(* IEC 61131-3 sources: SRCI_CLIENT_PLC/RobotLibrary/Library/Enumerations/Level, 5 files *)

(* ---- LogLevel.st ---- *)
{attribute 'qualified_only'}
// -------------------------------------------------------------------------
//  SRCI Robot Library
// -------------------------------------------------------------------------
//
//  Object:      LogLevel
//  Author:      Thorsten Brach
//  Date:        2024-06-01
//
//  Description:
//
//
//  Copyright:
//    (C) 2024 Thorsten Brach. All rights reserved
//             Licensed under the MIT License.
//
//  Disclaimer:
//    This project is provided without any guarantee and can be used for
//    private and commercial purposes. Any use is at the user’s
//    own risk and responsibility.
//
// -------------------------------------------------------------------------
// ST-FIX W02: no attribute 'to_string' - LogLevel is an alias of Severity, the attribute is only valid for enumerations
TYPE LogLevel : Severity; END_TYPE

(* ---- LogLevelEnum.st ---- *)
TYPE LogLevelEnum : LogLevel; END_TYPE

(* ---- MessageLevel.st ---- *)
{attribute 'qualified_only'}
{attribute 'to_string'}
// -------------------------------------------------------------------------
//  SRCI Robot Library
// -------------------------------------------------------------------------
//
//  Object:      MessageLevel
//  Author:      Thorsten Brach
//  Date:        2024-06-01
//
//  Description:
//
//
//  Copyright:
//    (C) 2024 Thorsten Brach. All rights reserved
//             Licensed under the MIT License.
//
//  Disclaimer:
//    This project is provided without any guarantee and can be used for
//    private and commercial purposes. Any use is at the user’s
//    own risk and responsibility.
//
// -------------------------------------------------------------------------
TYPE MessageLevel :
(
  /// Debugging messages, Informative messages, Warning messages, Error messages, Fatal error messages
  DEBUG := 4,
  /// Informative messages, Warning messages, Error messages, Fatal error messages
  INFO := 5,
  /// Warning messages, Error messages, Fatal error messages
  WARNING := 20,
  /// Error messages, Fatal error messages
  ERROR := 28
)USINT;
END_TYPE

(* ---- MessageLevelEnum.st ---- *)
TYPE MessageLevelEnum : MessageLevel; END_TYPE

(* ---- PriorityLevel.st ---- *)
{attribute 'qualified_only'}
{attribute 'to_string'}
// -------------------------------------------------------------------------
//  SRCI Robot Library
// -------------------------------------------------------------------------
//
//  Object:      PriorityLevel
//  Author:      Thorsten Brach
//  Date:        2024-06-01
//
//  Description:
//
//
//  Copyright:
//    (C) 2024 Thorsten Brach. All rights reserved
//             Licensed under the MIT License.
//
//  Disclaimer:
//    This project is provided without any guarantee and can be used for
//    private and commercial purposes. Any use is at the user’s
//    own risk and responsibility.
//
// -------------------------------------------------------------------------
TYPE PriorityLevel :
(
  /// priority level is very high
  VERY_HIGH := 1,
  /// priority level is high
  HIGH := 2,
  /// priority level is normal
  NORMAL := 3,
  /// priority level is low
  LOW := 4
)BYTE;
END_TYPE
